Staubli VAL3: cycle_Unhold.pgx

program cycle_Unhold()
begin
  //cycle进程:unholding
  rs:_nOmacStat=2
  //enable power
  if !isPowered()
    enablePower()
    watch(isPowered(),2)
  endIf
  restartMove()
  //cycle进程:running
  rs:_nOmacStat=3
  logMsg("当前处于生产状态 "+toString(".2",clock()))
  rs:_sRobotStatus="当前处于生产状态"
end
